TYPE ST_BhElFlow :
STRUCT
    eFlowUnit	:	E_BHElFlowUnit;

    {attribute 'pytmc' := '
        pv: Unit
        io: i
     '}
    i_sUnit			AT %I*	:	STRING;

    i_udiUnit	:	UDINT;

    {attribute 'pytmc' := '
        pv: Flow
        io: i
     '}
    i_rFlow			AT %I*	:	REAL;

    {attribute 'pytmc' := '
        pv: Setpoint
        io: o
     '}
    q_rSetpoint 	AT %Q*	:	REAL;

END_STRUCT
END_TYPE

(* stored: Version 1.1.0.1, ProductVersion 3.1.4022.18
   DUT ST_BhElFlow: Id {aa56882c-6739-4583-9306-a6edfd4b5ed1} *)
